(* IEC 61131-3 sources: daoli-st-library/DL_Process (part 6) *)

(* ---- FB_DL_ReactorStepCtrl.st ---- *)
(*==============================================================================
 * 组件名称 (Component)  : FB_DL_ReactorStepCtrl
 * 所属子库 (Sublibrary) : DL_Process
 * 前缀     (Prefix)     : FB_DL_
 * 当前版本 (Version)    : 1.0.1
 * 兼容性   (Platform)   : CODESYS 3.5 / TwinCAT 3 / 汇川 InoProShop / Schneider
 *                         Machine Expert；纯 IEC 61131-3（第 3 版），
 *                         仅依赖标准库 TON / R_TRIG / ABS / MAX / MIN 与库内
 *                         FB_DL_RampGenerator（IN-OUT 注入消费，斜坡不内联），
 *                         零厂商方言
 * 作者     (Author)     : 道莅代码库 · PLC编程专家（R31）
 * 开源溯源 (Origin)     : 反应釜工步顺控公开工艺语义（行业池）与 ISA-88 相
 *                         语义公开框架（暂停在步骤边界生效、恢复不重头，
 *                         主源记 T2-8），道莅 clean-room 防御性实现，
 *                         未复制任何外部源码行
 * 功能描述 (Function)   : 反应釜四工步顺控件：升温 → 保温 → 滴加 → 冷却。
 *                         温度设定经库内 FB_DL_RampGenerator 斜坡给出
 *                         （IN-OUT 注入，配方斜率单位 摄氏度每分钟 换算为
 *                         斜坡件的 摄氏度每秒 后下发）；滴加相以 bFeedAck
 *                         为终点带步超时；超温/超压独立监视层与顺控层
 *                         分离；暂停（bHold）在当前工步边界生效、恢复
 *                         不重头。不内联 PID（上层闭环外置）。
 * 复用清单 (Reuse)      : FB_DL_RampGenerator（斜坡设定，IN-OUT 注入）；
 *                         ISA-88 相语义（行为定义，零代码复制）。
 * 状态机   (States)     : eIdle/eHeat/eSoak/eFeed/eCool/eDone/ePaused/eFault，
 *                         CASE 带 ELSE 锁安全侧（fTSet 回零、停滴加）。
 * 码位     (Codes)      : 16#0005_00A8 信息级：配方域非法拒启动、配方钳位、
 *                                      暂停挂起提示（不置 bError）
 *                         16#0005_00A9 故障级：超温（独立监视层，锁存）
 *                         16#0005_00AA 故障级：超压（独立监视层，锁存）
 *                         16#0005_00AB 故障级：工步超时（滴加反馈缺失）
 *                         16#0005_00AC 故障级：状态非法（ELSE 兜底，锁存）
 * 边界防错 (Boundary)   : 1 配方域校验先于启动（斜率不大于零/温带倒置拒启动）；
 *                         2 bHold 仅在工步边界转暂停态，恢复续走原工步；
 *                         3 TON/R_TRIG 实例每拍无条件刷新；
 *                         4 CASE 带 ELSE 锁安全侧；
 *                         5 故障锁存可达解除路径：中止沿复归待机；
 *                         6 超温/超压监视独立于顺控相，任一相均生效。
 * 修订历史 (Revision)   : 2026-11-18 v1.0.0 首版入库（R31 · 阶段三 · 序 14）
 *                         2026-11-18 v1.0.1 R31 终审修复：中止/故障释放路径
 *                         补清 bError 与 uErrorId，消除释放后故障标志粘滞
 *==============================================================================*)

(*------------------------------------------------------------------------------
 * 结构体: ST_DL_ReactorRecipe（归属本功能块，同文件发布，全库唯一属主）
 *----------------------------------------------------------------------------*)
TYPE ST_DL_ReactorRecipe :
STRUCT
    fRampUp   : REAL := 2.0;    // 升温斜率 [摄氏度每分钟]，须大于 0 / Heat-up rate [degC per min], > 0
    fRampDown : REAL := 3.0;    // 降温斜率 [摄氏度每分钟]，须大于 0 / Cool-down rate [degC per min], > 0
    fSoakLo   : REAL := 80.0;   // 保温温带下限 [摄氏度] / Soak band lower [degC]
    fSoakHi   : REAL := 85.0;   // 保温温带上限 [摄氏度]，须高于下限 / Soak band upper [degC], above lower
    fFeedMl   : REAL := 50.0;   // 滴加量 [毫升] / Feed amount [mL]
    fCoolTgt  : REAL := 40.0;   // 冷却目标温度 [摄氏度] / Cool target temperature [degC]
END_STRUCT
END_TYPE

(*------------------------------------------------------------------------------
 * 枚举: E_DL_ReactorStep（归属本功能块，同文件发布，全库唯一属主）
 *----------------------------------------------------------------------------*)
TYPE E_DL_ReactorStep :
(
    eIdle   := 0,     // 待机：等待启动 / Idle, waiting for start
    eHeat   := 10,    // 升温工步：斜坡逼近温带 / Heat step, ramp to band
    eSoak   := 20,    // 保温工步：温带保持计时 / Soak step, hold band with timing
    eFeed   := 30,    // 滴加工步：等滴加反馈 / Feed step, wait feed acknowledgement
    eCool   := 40,    // 冷却工步：斜坡降到目标 / Cool step, ramp to target
    eDone   := 50,    // 完成：单拍脉冲后回待机 / Done, one-scan pulse then idle
    ePaused := 60,    // 暂停挂起：工步边界生效 / Paused, effective at step boundary
    eFault  := 99     // 故障：锁定等待中止复位 / Fault, latched until abort reset
);
END_TYPE

(*==============================================================================
 * 功能块: FB_DL_ReactorStepCtrl
 * 调用约定: 每个扫描周期无条件调用一次；ioRamp 为调用方持有的斜坡实例
 *           （IN-OUT 注入），本件驱动其引脚并读取其输出。
 *==============================================================================*)
FUNCTION_BLOCK FB_DL_ReactorStepCtrl
VAR_INPUT
    bStart   : BOOL := FALSE;         // 启动沿（待机且配方合法时受理）/ Start edge, accepted in idle with legal recipe
    bHold    : BOOL := FALSE;         // 暂停请求，工步边界生效 / Hold request, effective at step boundary
    bAbort   : BOOL := FALSE;         // 中止沿：任意态安全退出 / Abort edge, safe exit from any state
    fTNow    : REAL := 25.0;          // 釜温实测 [摄氏度] / Reactor temperature [degC]
    fPNow    : REAL := 101.0;         // 釜压实测 [千帕] / Reactor pressure [kPa]
    fPLimMax : REAL := 300.0;         // 超压监视限 [千帕]（可增引脚）/ Overpressure limit [kPa], added pin
    stRecipe : ST_DL_ReactorRecipe;   // 配方注入 / Recipe injected
    bFeedAck : BOOL := FALSE;         // 滴加完成反馈 / Feed acknowledgement feedback
    tSoak    : TIME := T#600S;        // 保温时长 [毫秒]（可增引脚）/ Soak duration [ms], added pin
    tFeedMax : TIME := T#600S;        // 滴加步超时 [毫秒]（可增引脚）/ Feed step timeout [ms], added pin
END_VAR
VAR_IN_OUT
    ioRamp   : FB_DL_RampGenerator;   // 斜坡发生器实例注入（库内复用）/ Ramp generator instance injected
END_VAR
VAR_OUTPUT
    eStep    : E_DL_ReactorStep;      // 当前工步 / Current step
    fTSet    : REAL;                  // 温度设定 [摄氏度]（斜坡输出）/ Temperature setpoint [degC]
    bFeedReq : BOOL;                  // 滴加请求 / Feed request
    bDone    : BOOL;                  // 全工步完成单拍脉冲（R27）/ All steps done one-scan pulse
    bError   : BOOL;                  // 故障标志，与故障级码配对（R45）/ Fault flag paired with fault codes
    uErrorId : UDINT;                 // 错误码，0 = 无错 / Error code, 0 = none
END_VAR
VAR
    rTrigStart: R_TRIG;               // 启动沿检测，每拍无条件刷新 / Start edge detector, refreshed every scan
    rTrigAbort: R_TRIG;               // 中止沿检测，每拍无条件刷新 / Abort edge detector, refreshed every scan
    tonSoak   : TON;                  // 保温计时，每拍无条件刷新 / Soak timer, refreshed every scan
    tonStep   : TON;                  // 步超时计时，每拍无条件刷新 / Step timeout timer, refreshed every scan
    bStepRst  : BOOL;                 // 步切换拍单拍断超时输入 / One-scan timeout break on step change
    eStatePrev: E_DL_ReactorStep;     // 上一拍步快照 / Previous step snapshot
    eResume   : E_DL_ReactorStep;     // 暂停前工步（恢复不重头）/ Step before pause, resume without restart
    bRcpOk    : BOOL;                 // 配方域合法标志 / Recipe legality flag
    bTValid   : BOOL;                 // 温度输入有效 / Temperature input validity
    bPValid   : BOOL;                 // 压力输入有效 / Pressure input validity
    bOverT    : BOOL;                 // 超温判定 / Over-temperature verdict
    bOverP    : BOOL;                 // 超压判定 / Over-pressure verdict
    uCodeLatch: UDINT;                // 故障级锁存码 / Latched fault code
    bInit     : BOOL := TRUE;         // 首扫标志 / First-scan flag
END_VAR
VAR CONSTANT
    DL_RSC_FIN   : REAL := 1.0E30;    // REAL 有限幅值判界 / REAL finiteness magnitude bound
    DL_RSC_OTMAR : REAL := 10.0;      // 超温监视裕度 [摄氏度] / Over-temp monitor margin [degC]
    DL_RSC_MIN2S : REAL := 60.0;      // 每分钟到每秒换算系数 / Per-min to per-sec factor
END_VAR

// ---- 段 1｜边沿与定时器实例无条件周期刷新（红线：禁入条件分支）----------------
rTrigStart(CLK := bStart);                            // 启动沿检测 / Start edge detection
rTrigAbort(CLK := bAbort);                            // 中止沿检测 / Abort edge detection
tonSoak(IN := (eStep = eSoak) AND (NOT bHold), PT := tSoak); // 保温计时，暂停断输入 / Soak timing, broken on hold
tonStep(IN := (eStep = eFeed) AND (NOT bStepRst), PT := tFeedMax); // 滴加超时按步断输入 / Feed timeout per step

// ---- 段 2｜步切换检测 ------------------------------------------------------------
bStepRst := (eStep <> eStatePrev) OR bInit;           // 步变化即断输入 / Step change breaks timing
eStatePrev := eStep;                                  // 快照留痕 / Snapshot previous step
bInit := FALSE;                                       // 清首扫标志 / Clear first-scan flag

// ---- 段 3｜输入有效性与独立监视层判定（与顺控相分离）------------------------------
bTValid := (fTNow = fTNow) AND (ABS(fTNow) < DL_RSC_FIN);   // 温度有限 / Temperature finite
bPValid := (fPNow = fPNow) AND (ABS(fPNow) < DL_RSC_FIN);   // 压力有限 / Pressure finite
bOverT  := bTValid AND (eStep <> eIdle) AND (fTNow > stRecipe.fSoakHi + DL_RSC_OTMAR); // 超温：带外裕度判 / Over-temp beyond margin
bOverP  := bPValid AND (eStep <> eIdle) AND (fPNow > fPLimMax); // 超压独立判 / Over-pressure independent
IF bOverT THEN
    uCodeLatch := 16#0005_00A9;                       // 码位：超温 / Code: over temperature
END_IF
IF bOverP THEN
    uCodeLatch := 16#0005_00AA;                       // 码位：超压 / Code: over pressure
END_IF
IF bOverT OR bOverP THEN
    eStep := eFault;                                  // 监视层直接锁故障 / Monitor layer latches fault directly
END_IF

// ---- 段 4｜中止沿统一入口：停滴加、温度设定回零、复归待机 ------------------------
IF rTrigAbort.Q THEN
    eStep := eIdle;                                   // 中止复归待机 / Abort returns to idle
    bFeedReq := FALSE;                                // 停滴加请求 / Stop feed request
    bError := FALSE;                                  // 中止含故障态释放路径，清故障标志（R28 终审）/ Abort is fault release path, clears flag
    uErrorId := 16#0000_0000;                         // 中止清错误码防粘滞（R28 终审）/ Abort clears error code against stickiness
END_IF

// ---- 段 5｜状态机（CASE 带 ELSE 锁安全侧：fTSet 回零、停滴加）---------------------
CASE eStep OF
    eIdle:
        fTSet := 0.0;                                 // 待机设定回零（安全侧）/ Idle setpoint zero, safe side
        bFeedReq := FALSE;                            // 待机停滴加 / Idle stops feed
        bDone := FALSE;                               // 清完成脉冲 / Clear done pulse
        ioRamp(bEnable := FALSE, bTrack := TRUE, fTrackValue := fTNow); // 斜坡跟踪实测免扰动 / Ramp tracks actual
        IF rTrigStart.Q THEN
            bRcpOk := (stRecipe.fRampUp > 0.0) AND (stRecipe.fRampDown > 0.0)
                  AND (stRecipe.fSoakLo < stRecipe.fSoakHi)
                  AND (stRecipe.fFeedMl >= 0.0) AND (stRecipe.fCoolTgt < stRecipe.fSoakLo)
                  AND (stRecipe.fRampUp < DL_RSC_FIN) AND (stRecipe.fRampDown < DL_RSC_FIN); // 配方域校验先于启动 / Recipe check before start
            IF bRcpOk THEN
                eStep := eHeat;                       // 配方合法进升温 / Legal recipe, to heat
            ELSE
                uErrorId := 16#0005_00A8;             // 信息级：配方非法拒启动 / Info: illegal recipe, start rejected
            END_IF
        END_IF
    eHeat:
        bFeedReq := FALSE;                            // 升温停滴加 / Heat stops feed
        ioRamp(bEnable := TRUE, fTarget := stRecipe.fSoakHi,
               fRateUp := stRecipe.fRampUp / DL_RSC_MIN2S,
               fRateDown := stRecipe.fRampDown / DL_RSC_MIN2S,
               bHold := FALSE);                       // 斜坡下发，配方斜率换算每秒 / Ramp driven, rate per second
        fTSet := ioRamp.fOut;                         // 温度设定取斜坡输出 / Setpoint from ramp output
        IF ioRamp.bDone AND bTValid AND (fTNow >= stRecipe.fSoakLo) THEN
            eStep := eSoak;                           // 到带复验后转保温（R42）/ Recheck then to soak
        END_IF
        IF bHold AND ioRamp.bDone THEN
            eResume := eSoak;                         // 边界暂停登记续点（ISA-88）/ Boundary pause books resume step
            eStep := ePaused;                         // 转暂停挂起 / To paused
        END_IF
    eSoak:
        bFeedReq := FALSE;                            // 保温停滴加 / Soak stops feed
        ioRamp(bEnable := TRUE, fTarget := stRecipe.fSoakHi,
               fRateUp := stRecipe.fRampUp / DL_RSC_MIN2S,
               fRateDown := stRecipe.fRampDown / DL_RSC_MIN2S,
               bHold := FALSE);                       // 保温维持带顶设定 / Soak holds band top
        fTSet := ioRamp.fOut;                         // 温度设定取斜坡输出 / Setpoint from ramp output
        IF tonSoak.Q THEN
            eStep := eFeed;                           // 保温满转滴加 / Soak elapsed, to feed
        END_IF
        IF bHold THEN
            eResume := eSoak;                         // 边界暂停登记续点 / Boundary pause books resume step
            eStep := ePaused;                         // 转暂停挂起 / To paused
        END_IF
    eFeed:
        bFeedReq := TRUE;                             // 滴加请求置位 / Feed request set
        fTSet := ioRamp.fOut;                         // 温度设定维持 / Setpoint maintained
        IF tonStep.Q THEN
            eStep := eFault;                          // 滴加反馈缺失锁故障（步超时）/ Feed ack missing, fault
            uCodeLatch := 16#0005_00AB;               // 码位：步超时/反馈缺失 / Code: step timeout
        ELSIF bFeedAck THEN
            eStep := eCool;                           // 滴加完成转冷却 / Feed done, to cool
        END_IF
    eCool:
        bFeedReq := FALSE;                            // 冷却停滴加 / Cool stops feed
        ioRamp(bEnable := TRUE, fTarget := stRecipe.fCoolTgt,
               fRateUp := stRecipe.fRampUp / DL_RSC_MIN2S,
               fRateDown := stRecipe.fRampDown / DL_RSC_MIN2S,
               bHold := FALSE);                       // 斜坡降到冷却目标 / Ramp down to cool target
        fTSet := ioRamp.fOut;                         // 温度设定取斜坡输出 / Setpoint from ramp output
        IF ioRamp.bDone AND bTValid AND (fTNow <= stRecipe.fCoolTgt + 1.0) THEN
            eStep := eDone;                           // 到目标复验后转完成（R42）/ Recheck then to done
        END_IF
        IF bHold AND ioRamp.bDone THEN
            eResume := eDone;                         // 边界暂停登记续点 / Boundary pause books resume step
            eStep := ePaused;                         // 转暂停挂起 / To paused
        END_IF
    eDone:
        fTSet := ioRamp.fOut;                         // 完成态维持设定 / Done maintains setpoint
        bFeedReq := FALSE;                            // 完成停滴加 / Done stops feed
        bDone := TRUE;                                // 完成单拍脉冲 / One-scan done pulse
        eStep := eIdle;                               // 下拍回待机 / Back to idle next scan
    ePaused:
        fTSet := ioRamp.fOut;                         // 暂停冻结设定（斜坡 bHold 语义由态承载）/ Pause freezes setpoint
        bFeedReq := FALSE;                            // 暂停停滴加 / Pause stops feed
        uErrorId := 16#0005_00A8;                     // 信息级：暂停挂起提示 / Info: paused notice
        IF (NOT bHold) AND (eResume <> ePaused) THEN
            eStep := eResume;                         // 恢复不重头续走原工步 / Resume without restart
        END_IF
    eFault:
        fTSet := 0.0;                                 // 故障安全侧设定回零 / Fault safe side setpoint zero
        bFeedReq := FALSE;                            // 故障停滴加 / Fault stops feed
        bDone := FALSE;                               // 故障清完成 / Fault clears done
        IF rTrigAbort.Q THEN
            eStep := eIdle;                           // 可达解除路径：中止沿复归 / Reachable release: abort edge
            uCodeLatch := 16#0000_0000;               // 清锁存码 / Clear latched code
            bError := FALSE;                          // 释放同步清故障标志（R28 终审）/ Release clears fault flag
            uErrorId := 16#0000_0000;                 // 释放同步清错误码 / Release clears error code
        END_IF
    ELSE
        eStep := eFault;                              // 非法状态兜底 / Illegal state fallback
        uCodeLatch := 16#0005_00AC;                   // 码位：状态非法 / Code: illegal state
        fTSet := 0.0;                                 // 兜底设定回零（安全侧）/ Fallback setpoint zero
        bFeedReq := FALSE;                            // 兜底停滴加 / Fallback stops feed
END_CASE

// ---- 段 6｜错误码装配：故障锁存回放优先，信息级居次 ------------------------------
IF eStep = eFault THEN
    bError   := TRUE;                                 // 故障标志配对（R45）/ Fault flag paired
    uErrorId := uCodeLatch;                           // 故障码锁存回放 / Latched fault code replayed
END_IF
END_FUNCTION_BLOCK

(* ---- FB_DL_ReworkLotGate.st ---- *)
(*
  ==================================================================
  组件名 Component  : FB_DL_ReworkLotGate
  分类   Category   : DL_Process
  前缀   Naming     : FB_DL_ ｜ b/n/u/f/t/e/st 类型前缀制（R265）
  码位   Code ID    : 16#0006_3036（故障级：越权放行锁存）｜ 16#0006_3037
                      （信息级：放行计数饱和钳位）
  版本   Version    : 1.0.1
  变更   CHANGELOG  : v1.0.1 eReleased 放行相单拍回迁
  复杂度 Complexity  : 中
  功能   Purpose    : 返工批拦截闸：返工标记登记期拦截放行指令，复检合格才
                      放行并计数；返工登记期未复检合格的放行指令判「越权
                      放行」并锁存故障；供批次放行合规审计与质量门禁使用。
  开源溯源 Origin    : ISA-88 批次相状态模型（公开条款，R12 沿用）+ PackML
                      纪律次源（T2-7 / T2-8）：仅借「批次相语义」状态命名
                      组织方式；返工闸逻辑完全自研，零代码复制。
  许可证 License    : MIT
  参考   Reference  : IEC 61131-3:2013 §6.6 状态机 / R_TRIG 语义；ISA-88
                      批次相状态公开条款（借语义，不抄文）
  平台   Platform   : 纯 IEC 61131-3（R_TRIG / ENUM+CASE / 四则），三平台通用
  依赖   Depends    : 仅 Standard.library（R_TRIG 属标准件）
  分工声明 Split     : FB_DL_BatchPhaseTrack（批次相跟踪）/ FB_DL_HoldResumeSeq
                      （保持恢复顺控）与本件互引；本件只管「返工标记 → 放行
                      合规」单门禁，不做批次全程跟踪（R216）。
  归属 Ownership     : E_DL_ReworkGatePhase 属主为本文件（全库唯一定义，R264）；
                      引用件只引用不重声明。
  ------------------------------------------------------------------
  边界 Boundary     :
                      一 组态口径（定稿，R90 反证句见码表）：nQuotaMax < 1
                         按「钳位接管为 1」静默接管——上限为 1 的闸仍有
                         完整拦截语义（登记 + 复检合格才放行 + 计数），
                         功能不静默丢失，非永假防御；不为此另立故障码
                         （组态缺省出口与正常运行出口完全同形：闸照常
                         工作、计数照常推进，无任何输出可区分该场景）；
                         3036 专用于越权放行锁存；
                      二 状态机 ENUM + CASE 必带 ELSE（非法态兜底落 eFault +
                         锁存 3036，禁静默）；本拍合法事件（复检合格沿 /
                         登记撤除）优先于越权判据（R275 同拍竞态）；
                      三 越权放行判据（锁存回放，R152）：返工登记电平 +
                         放行指令 + 复检未合格 → 锁存 3036 + bError；
                         锁存解除式（可达自证）：bResetCmd 上升沿清锁存
                         回 eIdle（输入引脚恒可达，无「置位即永久」路径）；
                      四 合规放行计数：放行沿（rtRelease R_TRIG，段 0 无条件
                         刷新）+ 复检合格 + 未锁存才计数；计数达 nQuotaMax
                         饱和钳位 + 信息级 3037（不置 bError，闸功能不受
                         影响，钳位为审计口径不是功能门槛）；
                      五 bEnable = FALSE 的语义写死（FB33-4 声明行）：强制
                         eIdle + 双出口复位（不 faults，使能断开 ≠ 合规故障）；
                      六 首拍 _bInit 全量初始化；无浮点量、无除法、无定时器
                         （纯电平 / 沿 / 计数语义）；无全局、无外部变量、
                         无物理地址。
  错误码 Codes      :
    16#0006_3036【故障级】越权放行（返工登记期放行指令且复检未合格）或非法
                         状态拦截（ELSE 兜底），锁存回放至复位沿
    16#0006_3037【信息级】放行计数已达 nQuotaMax 饱和钳位（不置 bError）
  码位反证 Note     :
    3036 与 3037 不可合并：3036 锁存 + bValid = FALSE + bError = TRUE，
    3037 不锁存 + bValid = TRUE + bError = FALSE，bValid / bError 双通道
    可唯一区分，按 R90 分立；「登记撤除瞬间的放行沿」与「越权」由同拍
    事件优先序区分（边界二），不需第三码。
  验收 Acceptance   :
    算法已证（脚本）：未跑 ｜ 编译器已证（三平台）：未跑
    V1 无登记 + 放行沿 → nReleased + 1、bReleaseAllow（正常批口径）
    V2 登记 + 复检合格 + 放行沿 → 计数 + 1（返工批合规放行）
    V3 登记 + 复检未合格 + 放行指令 → 锁存 3036 + bError
    V4 锁存态 bResetCmd 上升沿 → 解锁回 eIdle（锁存解除可达向量）
    V5 nQuotaMax = 3、放行 4 次 → nReleased 钳 3 + 码 3037
       （bError = FALSE，闸功能照常）
    V6 nQuotaMax = 0 → 钳位接管为 1（边界一定稿口径，功能不静默丢失）
    V7 失能 → eIdle + 双出口复位（不 faults）
    V8 非法枚举态（强改 eState）→ ELSE 兜底落 eFault + 3036
  修订记录 Revision  :
    2026-11-21  v1.0.0  R64 首版（批 3 · 序号 9，ISA-88 / PackML 纪律次源 + 自研）
    2026-11-22  v1.0.1  R65 点修（eReleased 回迁，R64 终审项）：v1.0.0 放行相
                        在 bReleaseCmd 持续保持且无再登记时停留该相不回迁，
                        下批次无法进入；v1.0.1 改放行相为单拍驻留相——完成后
                        无条件回迁待判 / 空闲相 eIdle；回迁清理声明：本件无
                        放行锁存与批次暂存变量（rtRelease 为自清沿实例，
                        Q 单拍自灭；nReleased 为审计台账不属暂存，复位沿亦
                        不清，边界四口径），回迁即天然清零，无需额外清零动作；
                        登记电平若仍生效，由 eIdle 相在下一拍重新迁入拦截相
                        （合法重入，rtRelease 沿不自触发，计数不受影响）
  ==================================================================
*)
TYPE E_DL_ReworkGatePhase :
(
    eIdle       := 0,  // 待机：无返工登记 / idle, no rework registered
    eReworkHold := 10, // 返工拦截：登记生效，等复检合格 / the rework hold, waiting for the recheck pass
    eReleased   := 20, // 放行：合规放行相（登记撤除或复检合格放行后驻留一拍语义由调用方承接）/ the released phase
    eFault      := 30  // 锁存故障：越权放行或非法态，复位沿解除 / a latched fault released by the reset edge
);
END_TYPE

FUNCTION_BLOCK FB_DL_ReworkLotGate
VAR_INPUT
    bEnable      : BOOL := TRUE;  // 使能，FALSE 时强制 eIdle + 双出口复位（边界五）/ the enable, false forces the idle and resets both outlets
    bLotRework   : BOOL := FALSE; // 返工标记登记电平 [-]（来自批次履历）/ the rework registration level from the lot history
    bRecheckPass : BOOL := FALSE; // 复检合格电平 [-] / the recheck pass level
    bReleaseCmd  : BOOL := FALSE; // 放行指令电平 [-] / the release command level
    bResetCmd    : BOOL := FALSE; // 故障复位电平，上升沿清锁存回 eIdle（边界三解除式）/ the fault reset level, its rising edge releases the latch
    nQuotaMax    : DINT  := 16;   // 放行计数饱和上限 [个]，须 ≥ 1，< 1 钳位接管为 1（边界一定稿）/ the release count ceiling, at least one, clamped when below
END_VAR
VAR_OUTPUT
    bReleaseAllow : BOOL := FALSE;           // 放行许可电平 [-]（锁存 / 失能强制 FALSE）/ the release permission forced false on a latch or disable
    bReworkHold   : BOOL := FALSE;           // 返工拦截中指示 [-] / the rework hold indicator
    nReleased     : DINT  := 0;              // 合规放行计数 [个]（饱和口径）/ the compliant release count saturated
    eState        : E_DL_ReworkGatePhase;    // 状态机出口 [状态] / the state machine outlet
    bValid        : BOOL := FALSE;           // 判据可用 [-] / the criteria are usable
    eErr          : UDINT := 16#0000_0000;   // 错误码，0 = 正常 / the error code, zero is ok
    bError        : BOOL := FALSE;           // 故障标志（故障级码同拍置位，R45 配对）/ the fault flag raised with a fault level code
END_VAR
VAR
    _bInit      : BOOL := FALSE;  // 首拍初始化标志（R310 / FB50-2）/ the first scan flag
    _eState     : E_DL_ReworkGatePhase := E_DL_ReworkGatePhase.eIdle; // 内部状态寄存器 / the internal state register
    _bFaultLatch: BOOL := FALSE;  // 故障锁存副本（仅复位沿清除）/ the fault latch copy
    _uLatch     : UDINT := 16#0000_0000; // 故障码锁存 [码]（复位沿清除，FB33-1）/ the latched fault code cleared by the reset edge
    _nReleased  : DINT  := 0;     // 计数内部副本 [个]（饱和钳位口径）/ the internal count copy saturated
    _nQuotaUse  : DINT  := 1;     // 上限接管量 [个]（< 1 钳位为 1，边界一）/ the ceiling taken over clamped to one
    _bCountSat  : BOOL := FALSE;  // 计数饱和标记（单拍信息位，段 6 映射）/ the count saturation flag of this scan
    rtReset     : R_TRIG;         // 复位沿实例，段 0 无条件刷新（R7）/ the reset edge instance refreshed unconditionally
    rtRelease   : R_TRIG;         // 合规放行沿实例，段 0 无条件刷新 / the compliant release edge instance refreshed unconditionally
END_VAR  // R64 结构补齐：VAR 段缺失的 END_VAR（门禁机械修复）
VAR CONSTANT
    DL_RLG_ZEROI: DINT  := 0;  // 整型零常量 [个] / the integer zero constant
    DL_RLG_ONEI : DINT  := 1;  // 整型一常量 [个] / the integer one constant
    DL_RLG_ZEROU: UDINT := 16#0000_0000; // 码零常量 / the code zero constant
END_VAR

// 段 0｜沿检测无条件周期刷新（禁入分支，R7）/ segment 0, the unconditional edge refresh
rtReset(CLK := bResetCmd); // 复位沿 / the reset edge
rtRelease(CLK := bReleaseCmd AND NOT _bFaultLatch AND bEnable
                 AND (NOT bLotRework OR bRecheckPass)); // 合规放行沿（登记撤除或复检合格的放行指令上升沿，R275 事件优先口径）/ the compliant release edge of the legal command

// 段 1｜首拍初始化与复位沿作用域（R310 / R311）/ segment 1, the first scan init and the reset edge scope
IF NOT _bInit THEN // 首拍一拍 / the first scan
    _bInit := TRUE; // 置首拍标志 / raise the first scan flag
    _eState := E_DL_ReworkGatePhase.eIdle; // 状态显式落空闲 / place the state to idle
    _bFaultLatch := FALSE; // 故障锁存显式清零 / clear the fault latch explicitly
    _uLatch := DL_RLG_ZEROU; // 码锁存显式清零 / clear the latched code explicitly
    _nReleased := DL_RLG_ZEROI; // 计数显式清零 [个] / clear the count explicitly
    _nQuotaUse := DL_RLG_ONEI; // 上限接管显式置一 [个] / preset the ceiling one explicitly
END_IF
IF rtReset.Q THEN // 复位沿（作用域声明：清锁存 + 迁相位，不清计数——计数是审计台账，R311）/ the reset edge with the declared scope, the audit count survives
    _bFaultLatch := FALSE; // 清故障锁存（唯一解除路径，边界三自证可达）/ clear the fault latch, the only release path
    _uLatch := DL_RLG_ZEROU; // 清码锁存 / clear the latched code
    _eState := E_DL_ReworkGatePhase.eIdle; // 迁回空闲 / back to idle
END_IF

// 段 2｜上限接管与计数饱和预置（边界一：nQuotaMax < 1 钳位接管为 1，功能不静默丢失）/ segment 2, the ceiling take over and the saturation preset
_nQuotaUse := nQuotaMax; // 上限接管 [个] / take the ceiling
IF _nQuotaUse < DL_RLG_ONEI THEN // 上限 < 1（组态缺省）/ the ceiling below one
    _nQuotaUse := DL_RLG_ONEI; // 钳位接管为 1（拦截闸仍有完整语义）/ clamp to one, the gate keeps its full semantics
END_IF
_bCountSat := FALSE; // 计数饱和标记预清零（单拍信息位，R256 统一出口预置）/ preset the saturation flag false

// 段 3｜失能分支：强制 eIdle + 双出口复位，不 faults（边界五声明行）/ segment 3, the disabled branch
IF NOT bEnable THEN // 失能 / disabled
    _eState := E_DL_ReworkGatePhase.eIdle; // 强制空闲 / force the idle
    _bFaultLatch := FALSE; // 锁存复位（使能断开 ≠ 合规故障）/ clear the latch
    _uLatch := DL_RLG_ZEROU; // 码锁存复位 / clear the code
    eState := _eState; // 状态出口 / the state outlet
    bReleaseAllow := FALSE; // 许可电平复位 / the permission resets
    bReworkHold := FALSE; // 拦截指示复位 / the hold indicator resets
    bValid := FALSE; // 失能即不可用 / the criteria are not usable while disabled
    bError := FALSE; // 失能不是故障 / a disabled device is not a fault
    eErr := DL_RLG_ZEROU; // 失能不发码 / no code is emitted while disabled
    RETURN; // 早退（计数不动，失能不清审计台账）/ early return, the audit count survives
END_IF

// 段 4｜主状态机（ENUM + CASE，ELSE 兜底；本拍事件优先于越权判据，R275）/ segment 4, the main machine, the event before the misuse verdict
CASE _eState OF
    E_DL_ReworkGatePhase.eIdle: // 空闲相 / the idle phase
        IF bLotRework THEN // 返工登记生效 / the rework registration is active
            _eState := E_DL_ReworkGatePhase.eReworkHold; // 迁入拦截相 / enter the hold phase
        END_IF
    E_DL_ReworkGatePhase.eReworkHold: // 返工拦截相（本拍合法事件优先：登记撤除或复检合格放行先消化，再消化越权判据，R275）/ the hold phase, the legal event before the misuse
        IF NOT bLotRework THEN // 事件优先：登记撤除 / the registration withdrawn, the event goes first
            _eState := E_DL_ReworkGatePhase.eIdle; // 回空闲 / back to idle
        ELSIF bRecheckPass AND bReleaseCmd THEN // 复检合格 + 放行指令（合规放行，边界四口径）/ the recheck passed with the release command
            _eState := E_DL_ReworkGatePhase.eReleased; // 迁入放行相 / enter the released phase
        ELSIF bReleaseCmd THEN // 越权判据：登记中放行且复检未合格（真实可达：操作员越过复检直接放令）/ the misuse path, reachable by the operator bypassing the recheck
            _bFaultLatch := TRUE; // 锁存故障 / latch the fault
            _uLatch := 16#0006_3036; // 故障级：越权放行 / fault grade, the unauthorized release
            bError := TRUE; // 同拍置故障标志（R45 配对，段 6 故障分支沿用）/ raise the fault flag on the same scan
        END_IF
    E_DL_ReworkGatePhase.eReleased: // 放行相（v1.0.1 改单拍驻留：完成后强制回迁空闲，R64 终审修复「eReleased 不回迁」）/ the released phase, single scan dwell with the forced return since v1.0.1
        _eState := E_DL_ReworkGatePhase.eIdle; // 放行相完成后无条件回迁待判 / 空闲相（下批次可正常进入；v1.0.0 在 bReleaseCmd 持续保持且无再登记时停留该相不回迁，为本次修复点）/ unconditional return to idle after the release completes
        // 回迁清理声明（v1.0.1）：本件无放行锁存与批次暂存变量——rtRelease 为自清沿实例（Q 单拍自灭），nReleased 为审计台账不属暂存（复位沿亦不清，边界四），回迁即天然清零，无额外清零动作 / no release latch or batch staging exists, the return clears naturally
    E_DL_ReworkGatePhase.eFault: // 锁存故障相（驻留，解除由段 1 复位沿承担）/ the fault phase dwelling, the release belongs to the reset edge
        ; // 驻留语义由注释表达（禁自赋值死语句，R261）/ the dwell is expressed by this comment without a dead statement
    ELSE // 非法枚举值拦截（边界二：落故障相并锁存，禁静默）/ the illegal enumeration guard
        _bFaultLatch := TRUE; // 锁存故障 / latch the fault
        _uLatch := 16#0006_3036; // 故障级：非法状态拦截（归入越权族一码，出口同形锁存回放，R90）/ fault grade, the illegal state under the latch family
        bError := TRUE; // 同拍置故障标志（R45 配对）/ raise the fault flag on the same scan
        _eState := E_DL_ReworkGatePhase.eFault; // 落故障相 / force the fault phase
END_CASE

// 段 5｜合规放行计数（边界四：沿 + 未锁存才计数；饱和钳位 + 信息级）/ segment 5, the compliant release counting with the saturation
IF rtRelease.Q AND (NOT _bFaultLatch) THEN // 合规放行沿且未锁存 / a compliant release edge without a latch
    IF _nReleased < _nQuotaUse THEN // 计数未达上限 / the count below the ceiling
        _nReleased := _nReleased + DL_RLG_ONEI; // 计数推进 [个] / advance the count
    ELSE // 计数已达上限：饱和钳位 + 信息级（闸功能不受影响，边界四）/ the count saturated with the info code, the gate unaffected
        _bCountSat := TRUE; // 置饱和标记（单拍信息位）/ raise the saturation flag
    END_IF
END_IF

// 段 6｜故障锁存迁移闸 + 统一出口（名实双出口同源，R191）/ segment 6, the latch gate and the unified outlet
IF _bFaultLatch AND (_eState <> E_DL_ReworkGatePhase.eFault) THEN // 已锁存但不在故障相 / latched outside the fault phase
    _eState := E_DL_ReworkGatePhase.eFault; // 迁入故障相 / enter the fault phase
END_IF
eState := _eState; // 状态出口 / the state outlet
bReleaseAllow := (NOT _bFaultLatch) AND bEnable
              AND ((NOT bLotRework) OR bRecheckPass); // 许可电平与判据同源派生（登记中须复检合格）/ the permission derived from the criteria
bReworkHold := (_eState = E_DL_ReworkGatePhase.eReworkHold); // 拦截指示与状态同源 / the hold indicator from the state
nReleased := _nReleased; // 计数出口 [个] / the count outlet
IF _bFaultLatch THEN // 故障锁存回放优先（不在故障相按当下输入重新推断，R152）/ the latched fault replays first
    bValid := FALSE; // 故障相不可用 / not usable in the fault phase
    bError := TRUE; // 故障位置位（R45 配对）/ raise the fault bit
    eErr := _uLatch; // 锁存码回放 / replay the latched code
ELSIF _bCountSat THEN // 计数饱和（信息级，单拍重算）/ the saturation, informational
    bValid := TRUE; // 闸功能照常可用 / the gate stays usable
    bError := FALSE; // 信息级不置故障标志（R285）/ keep the fault flag false
    eErr := 16#0006_3037; // 信息级：放行计数饱和钳位 / informational, the count saturated
ELSE // 无事件 / no event
    bValid := TRUE; // 判据可用 / the criteria are usable
    bError := FALSE; // 无故障 / no fault
    eErr := DL_RLG_ZEROU; // 正常 / ok
END_IF
END_FUNCTION_BLOCK

(* ---- FB_DL_RotaryIndexTable.st ---- *)
(*==============================================================================
 * 组件名称 (Component)  : FB_DL_RotaryIndexTable
 * 所属子库 (Sublibrary) : DL_Process
 * 当前版本 (Version)    : 1.0.0
 * 组件分类 (Category)   : 功能块（FUNCTION_BLOCK）· 工站模板 · 多工位分度盘调度
 * 兼容性 (Platform)     : CODESYS 3.5 / TwinCAT 3 / 汇川 InoProShop / Machine Expert；
 *                         仅依赖标准库（TON / R_TRIG / F_TRIG / LIMIT），分度请求
 *                         以布尔脉冲出口下发，块内不绑定任何电机或驱动库
 * 功能描述 (Function)   : 管理「分度请求 → 到位确认 → 稳定等待 → 工位工艺放行」的
 *                         节拍链；维护工位启用表与工艺号映射，支持空跑（清洗）模式
 *                         逐位走完，并对分度超时与到位信号抖动给出可诊断的故障码
 * 与既有件边界 (Scope)  : 料仓槽位台账（空 / 满 / 不合格）由料仓件承担，本块不管槽
 *                         位内容；连续输送积放由输送段件承担，本块管离散分度盘的节
 *                         拍与工位放行。三者拓扑互斥，语义不重叠
 * 状态机规模 (States)   : 五态最小子集（eIdle 0 / eDwell 10 / eIndexing 20 /
 *                         eSettling 30 / eFault 99）。eSettling 单独成态，用于隔离
 *                         「到位后抖动」的诊断窗口，避免把机械抖动混入分度超时计数
 * 关键算法 (Algorithm)  :
 *   ① 工位号合法性：nAtStation 须落在 1~生效工位数，越界即 02D2，不做猜测性修正
 *   ② 掩码构造：每拍由启用表重建，逐位置位（位累加器左移一位再或），不拼累计量，
 *      规避位宽边界；工位数上限 24，恒在安全域内
 *   ③ 停留计时：剩余停留时间由定时器已历时反算，空跑模式直接旁路计时
 *   ④ 空跑模式：工艺放行恒假，分度链照走，用于清洗与调试；不计循环数
 *   ⑤ 循环计数：分度回到 1 号位那一拍出单拍脉冲并累加，饱和防溢出
 *   ⑥ 抖动诊断：稳定窗内到位信号掉沿即判硬件问题，直接锁故障且不自动重试——自动
 *      重试会把机械松动掩盖成偶发超时，现场极难定位
 * 码位表 (Error codes)  :
 *   16#0005_01C2【信息级】工位数量越界已钳位至 2~24，不置故障位
 *   16#0005_02D0【故障级】分度超时（到位信号未在监控窗内建立）
 *   16#0005_02D1【故障级】到位信号抖动或丢失（稳定窗内掉沿）
 *   16#0005_02D2【故障级】工位号越界（机械到位反馈不可信）
 *   16#0005_02D3【故障级】非法状态兜底
 * R32 写入点次序审计 :
 *   nActiveStation  : ① 空跑 / 停机撤销时清 0（段 6、段 7）→ ② 停留与稳定段按到位
 *                     反馈刷新（eDwell / eSettling 各一处，同拍只可能命中一处）
 *   bStationReady   : 仅段 10 单点派生（由生效工位数、启用表、空跑模式三者与门），
 *                     状态机内不写，杜绝分支双写
 *   nRecipeAtStation: 仅段 10 单点派生（工艺号透传，越界给 0，不做校验）
 *   tDwellRemain    : 仅段 10 单点派生（由停留定时器已历时反算，钳位非负）
 *   _uErrorIdInt    : ① 首扫清（段 4）→ ② 分度超时（eIndexing）→ ③ 抖动（eSettling）
 *                     → ④ 工位号越界（eSettling）→ ⑤ 非法状态（ELSE）→ ⑥ 复位清
 *   _eState         : 每拍只在 CASE 分支出口单点写入；CASE 之外仅段 6 使能撤销一处
 * 设计偏离登记 (Deviations) :
 *   D1 增补 tCycle 引脚（默认 10 毫秒）：统计结构体内含累计运行时长，而块内无时间
 *      基准引脚则无法累加；按库内既有公约以任务扫描周期作基准，向后兼容（有默认
 *      值），不改变任何既有引脚语义
 *   D2 分度计数在「到位确认通过」拍累加，而非请求拍：超时未到位属失败分度，不应
 *      计入成功次数；与规格文字「分度次数」取成功口径一致
 * 验收向量 (Acceptance) :
 *   V1 掩码：工位数 8、前 5 个启用 → 掩码 16#0000_001F
 *   V2 工艺号透传：到位 3 号工位、3 号工艺号 27 → 作业工位 3、工艺号 27、放行为真
 *   V3 分度超时：监控窗 2 秒内到位信号未建立 → 码 02D0、故障态、故障位为真
 *   V4 空跑：工位数 4、空跑为真 → 逐位推进，4 拍后出循环脉冲，循环计数不增
 *   V5 抖动：到位后 50 毫秒内信号由真转假 → 码 02D1，无自动重试
 * 开源溯源 (Origin)     : 参考包装机械公开手册的工位 / 节拍语义组织与位掩码工位表
 *                         写法，只借分类与参数域；状态机、掩码重建、抖动诊断、码位
 *                         与引脚契约为本库独立设计，clean-room 不构成衍生作品
 * 红线自检 (Redline)    : R1 零全局表与外部变量引用、零物理地址记号 ✓｜R2 零占位符 ✓
 *                         R3 纯 IEC 61131-3 加标准库 ✓｜R4 数组先判界、除法防零、
 *                         时长反算钳非负 ✓｜R5 声明行中英双语同行注释 ✓｜R6 五成员逐
 *                         一有 CASE 标签且含 ELSE 兜底 ✓｜R7 三沿检测（启动 / 停止 /
 *                         复位）与到位双沿、三定时器全部在 CASE 之外无条件刷新 ✓
 * 修订历史 (Revision)   :
 *   2026-11-15  v1.0.0  首版入库（Round 11 · C 泳道 · 工站四件套之二）
 *============================================================================*)

(*------------------------------------------------------------------------------
 * 枚举: E_DL_IndexTableState（归属 FB_DL_RotaryIndexTable，同文件发布）
 *   五态，每个成员在主状态机中均有同名 CASE 标签（R31 完备性）
 *-----------------------------------------------------------------------------*)
TYPE E_DL_IndexTableState :
(
    eIdle     := 0,     // 待机：等启动沿，不发放行 / Idle, awaiting start, no permit
    eDwell    := 10,    // 停留：当前工位工艺放行窗 / Dwell, process permit window
    eIndexing := 20,    // 分度中：已出请求脉冲，等到位 / Indexing, waiting for in-position
    eSettling := 30,    // 稳定中：到位后去抖确认 / Settling, debounce after in-position
    eFault    := 99     // 故障锁存：仅复位沿可退 / Fault latched, only a reset edge leaves
);
END_TYPE

(*------------------------------------------------------------------------------
 * 结构体: ST_DL_IndexTableStat（归属 FB_DL_RotaryIndexTable）
 *   跨周期统计，由调用方持有，本块只累加，掉电保持由上层负责
 *-----------------------------------------------------------------------------*)
TYPE ST_DL_IndexTableStat :
STRUCT
    nIndexCount : UDINT;                    // 累计成功分度次数 [次] [Successful index counter]
    nCycleCount : UDINT;                    // 累计整圈循环数 [圈] [Full revolution counter]
    tRunTime    : TIME;                     // 累计运行时长 [毫秒] [Accumulated run time]
END_STRUCT
END_TYPE

FUNCTION_BLOCK FB_DL_RotaryIndexTable
VAR_INPUT
    bEnable          : BOOL;                            // 使能，FALSE 撤销分度请求并回待机 [Enable, withdraws request on FALSE]
    bStart           : BOOL;                            // 启动节拍循环，上升沿受理 [Start the cycle on a rising edge]
    bStop            : BOOL;                            // 完成当前工位后停止，上升沿受理 [Stop after current station, rising edge]
    bReset           : BOOL;                            // 复位故障，上升沿受理 [Reset fault on rising edge]
    nStationCount    : INT;                             // 工位总数 [个]，有效域 2~24 [Station count, 2..24]
    nAtStation       : INT;                             // 机械到位工位号 [1~工位数]，0 表示未定位 [Mechanical station number, 0 = not seated]
    bIndexInPos      : BOOL;                            // 分度到位开关信号 [-] [Indexer in-position switch]
    abStationEnable  : ARRAY[1..24] OF BOOL;            // 工位启用表，FALSE 视为空位 [Station enable table, FALSE = empty]
    anStationRecipe  : ARRAY[1..24] OF INT;             // 工位工艺号表，仅透传不校验 [-] [Per-station recipe number, pass-through]
    tDwellTime       : TIME := T#1S;                    // 每工位停留时间 [毫秒]，0 表示不停留 [Dwell per station]
    tSettleTime      : TIME := T#100MS;                 // 到位后稳定确认时间 [毫秒]，滤机械抖动 [Settling time after in-position]
    tIndexTimeout    : TIME := T#3S;                    // 分度超时 [毫秒]，0 表示不监控 [Indexing timeout]
    bDryRun          : BOOL;                            // 空跑（清洗）模式：忽略启用表逐位走完 [Dry-run mode, ignores enable table]
    tCycle           : TIME := T#10MS;                  // 任务扫描周期 [毫秒]，累计运行时长基准（偏离 D1）[Task cycle time, run-time base]
END_VAR
VAR_OUTPUT
    bIndexReq        : BOOL;                            // 分度请求，单拍脉冲 [-] [Index request, single-scan pulse]
    nActiveStation   : INT;                             // 当前作业工位号 [1~工位数]，0 表示无效 [Active station number, 0 = invalid]
    bStationReady    : BOOL;                            // 当前工位允许工艺动作 [-] [Station ready for process action]
    nRecipeAtStation : INT;                             // 当前工位工艺号，透传 [-] [Recipe number at active station]
    uStationMask     : DWORD;                           // 工位启用镜像，第 n 位对应第 n 工位 [Station enable mirror, bit n-1]
    bCycleDone       : BOOL;                            // 整圈走完单拍脉冲 [-] [Single pulse on full revolution]
    tDwellRemain     : TIME;                            // 当前工位剩余停留时间 [毫秒] [Remaining dwell time]
    eState           : E_DL_IndexTableState;            // 主状态机当前态 [-] [Current state]
    bError           : BOOL;                            // 故障锁存，需复位清除 [Latched fault]
    uErrorId         : UDINT;                           // 事件码或故障码，0 表示无 [Event or fault code]
END_VAR
VAR_IN_OUT
    stStat           : ST_DL_IndexTableStat;            // 跨周期统计，调用方持有 [Persistent statistics]
END_VAR
VAR
    _eState          : E_DL_IndexTableState := E_DL_IndexTableState.eIdle;  // 内部状态寄存器，唯一真值源 [Internal state register]
    _bInit           : BOOL := FALSE;                   // 首扫标志，初值 FALSE，判据 NOT _bInit [First-scan flag, R19 pattern]
    _bFaultLatch     : BOOL;                            // 故障级锁存，仅复位路径清 [Fault latch, reset path only]
    _uErrorIdInt     : UDINT;                           // 故障级码寄存 [Fault-level code register]
    _uInfoCode       : UDINT;                           // 本拍信息级码，每拍重算 [Transient info code]
    nStaEff          : INT;                             // 生效工位数，已钳位 [个] [Effective station count]
    nIdxVal          : INT;                             // 到位工位号（已判界）[号] [Validated station number]
    tDwellEff        : TIME;                            // 生效停留时间 [毫秒] [Effective dwell time]
    tSettleEff       : TIME;                            // 生效稳定时间 [毫秒] [Effective settling time]
    tIndexEff        : TIME;                            // 生效分度超时 [毫秒] [Effective index timeout]
    tCycleEff        : TIME;                            // 生效扫描周期 [毫秒] [Effective task cycle time]
    uMaskAcc         : UDINT;                           // 掩码累加器 [位域] [Mask accumulator]
    uBitAcc          : UDINT;                           // 位累加器，逐位左移 [位域] [Single-bit accumulator]
    nI               : INT;                             // 通用循环索引 [索引] [Loop index]
    bDwellIn         : BOOL;                            // 停留计时输入条件，先算后调 [Dwell timer input]
    bSettleIn        : BOOL;                            // 稳定计时输入条件，先算后调 [Settle timer input]
    bIndexIn         : BOOL;                            // 分度超时输入条件，先算后调 [Index timer input]
    bDwellDone       : BOOL;                            // 停留结束（含空跑旁路）[Dwell finished, dry-run bypassed]
    _bInPosDropped   : BOOL;                            // 分度中到位信号曾回落，兼容保持型开关 [In-position dropped during indexing]
    fbTrigStart      : R_TRIG;                          // 启动沿检测 [Start edge detector]
    fbTrigStop       : R_TRIG;                          // 停止沿检测 [Stop edge detector]
    fbTrigReset      : R_TRIG;                          // 复位沿检测 [Reset edge detector]
    fbTrigInPos      : R_TRIG;                          // 到位上升沿检测 [In-position rising edge]
    fbTrigInPosFall  : F_TRIG;                          // 到位下降沿检测，抖动诊断用 [In-position falling edge, jitter diagnosis]
    fbTmoDwell       : TON;                             // 停留计时 [Dwell timer]
    fbTmoSettle      : TON;                             // 稳定确认计时 [Settle timer]
    fbTmoIndex       : TON;                             // 分度超时 [Index timeout timer]
END_VAR
VAR CONSTANT
    DL_STATION_MAX   : INT := 24;                       // 工位上限 [个] [Max station count]
    DL_STATION_MIN   : INT := 2;                        // 工位下限 [个] [Min station count]
    DL_TMO_MAX       : TIME := T#120S;                  // 时长参数域上限 [毫秒] [Duration upper bound]
    DL_RUN_MAX       : TIME := T#500H;                 // 运行时长饱和上限 [毫秒] [Run time saturation limit]
    DL_COUNT_MAX     : UDINT := 16#FFFF_FFFE;           // 计数饱和上限 [次] [Counter saturation limit]
    DL_INFO_STA_CLAMP: UDINT := 16#0005_01C2;           // 01C2 工位数量越界已钳位【信息级】 [Info, station count clamped]
    DL_ERR_INDEX_TMO : UDINT := 16#0005_02D0;           // 02D0 分度超时【故障级】 [Fault, index timeout]
    DL_ERR_INPOS     : UDINT := 16#0005_02D1;           // 02D1 到位信号抖动或丢失【故障级】 [Fault, in-position lost]
    DL_ERR_STATION   : UDINT := 16#0005_02D2;           // 02D2 工位号越界【故障级】 [Fault, station out of range]
    DL_ERR_STATE     : UDINT := 16#0005_02D3;           // 02D3 非法状态兜底【故障级】 [Fault, illegal state]
END_VAR

// ==== 段 1｜单拍输出预清零（脉冲类出口每拍先清零，避免跨拍粘滞） / Single-scan pulse pre-clear, no sticky pulses
bIndexReq  := FALSE;                        // 分度请求先清零 [Index request pre-cleared]
bCycleDone := FALSE;                        // 整圈完成先清零 [Revolution pulse pre-cleared]
_uInfoCode := 16#0000_0000;                 // 信息级码每拍重算 [Info code recomputed]

// ==== 段 2｜参数钳位（工位数与三个时长，先钳位再进逻辑） / Parameter clamping before any logical use
nStaEff := nStationCount;                   // 工位数先取引脚值 [Station count from pin]
IF nStaEff < DL_STATION_MIN THEN
    nStaEff    := DL_STATION_MIN;           // 低于下限钳到 2 [Clamped to lower bound]
    _uInfoCode := DL_INFO_STA_CLAMP;        // 01C2 工位数量越界已钳位【信息级】 [Info, count clamped]
ELSIF nStaEff > DL_STATION_MAX THEN
    nStaEff    := DL_STATION_MAX;           // 高于上限钳到 24 [Clamped to upper bound]
    _uInfoCode := DL_INFO_STA_CLAMP;        // 01C2 工位数量越界已钳位【信息级】 [Info, count clamped]
END_IF

tDwellEff := tDwellTime;                    // 停留时间先取引脚值 [Dwell from pin]
IF tDwellEff > DL_TMO_MAX THEN
    tDwellEff := DL_TMO_MAX;                // 超上限钳位 [Clamped to upper bound]
ELSIF tDwellEff < T#0S THEN
    tDwellEff := T#0S;                      // 负值归零 [Negative clamped to zero]
END_IF

tSettleEff := tSettleTime;                  // 稳定时间先取引脚值 [Settle from pin]
IF tSettleEff > DL_TMO_MAX THEN
    tSettleEff := DL_TMO_MAX;               // 超上限钳位 [Clamped to upper bound]
ELSIF tSettleEff < T#0S THEN
    tSettleEff := T#0S;                     // 负值归零 [Negative clamped to zero]
END_IF

tIndexEff := tIndexTimeout;                 // 分度超时先取引脚值 [Index timeout from pin]
IF tIndexEff > DL_TMO_MAX THEN
    tIndexEff := DL_TMO_MAX;                // 超上限钳位 [Clamped to upper bound]
ELSIF tIndexEff <= T#0S THEN
    tIndexEff := T#0S;                      // 零表示不监控 [Zero means supervision disabled]
END_IF

tCycleEff := tCycle;                        // 扫描周期先取引脚值 [Task cycle from pin]
IF tCycleEff <= T#0S OR tCycleEff > T#10S THEN
    tCycleEff := T#10MS;                    // 异常值回默认 10 毫秒 [Fallback to 10 ms]
END_IF

// ==== 段 3｜沿与定时器无条件刷新（R7 红线：严禁置于 IF / CASE 分支内） / Unconditional refresh of edges and timers
fbTrigStart(CLK := bStart);                 // 启动沿 [Start edge]
fbTrigStop(CLK := bStop);                   // 停止沿 [Stop edge]
fbTrigReset(CLK := bReset);                 // 复位沿 [Reset edge]
fbTrigInPos(CLK := bIndexInPos);            // 到位上升沿 [In-position rising edge]
fbTrigInPosFall(CLK := bIndexInPos);        // 到位下降沿 [In-position falling edge]

IF _eState = E_DL_IndexTableState.eDwell THEN
    bDwellIn := TRUE;                       // 仅停留段计时 [Only during dwell]
ELSE
    bDwellIn := FALSE;                      // 其余段清零 [Cleared otherwise]
END_IF
fbTmoDwell(IN := bDwellIn, PT := tDwellEff);

IF _eState = E_DL_IndexTableState.eSettling THEN
    bSettleIn := TRUE;                      // 仅稳定段计时 [Only during settling]
ELSE
    bSettleIn := FALSE;                     // 其余段清零 [Cleared otherwise]
END_IF
fbTmoSettle(IN := bSettleIn, PT := tSettleEff);

IF (_eState = E_DL_IndexTableState.eIndexing) AND (tIndexEff > T#0S) THEN
    bIndexIn := TRUE;                       // 仅分度段且监控开启时计时 [Only while indexing with supervision on]
ELSE
    bIndexIn := FALSE;                      // 其余段清零 [Cleared otherwise]
END_IF
fbTmoIndex(IN := bIndexIn, PT := tIndexEff);

// ==== 段 4｜首扫初始化（R19 唯一合法范式：初值 FALSE，判据 NOT，同步后置 TRUE） / First-scan initialisation with the canonical R19 pattern
IF NOT _bInit THEN
    _eState          := E_DL_IndexTableState.eIdle;  // 状态回待机 [State to idle]
    _bInPosDropped   := FALSE;              // 到位回落标志复位 [Dropped flag reset]
    _bFaultLatch     := FALSE;              // 故障锁存清零 [Fault latch cleared]
    _uErrorIdInt     := 16#0000_0000;       // 故障码清零 [Fault code cleared]
    nActiveStation   := 0;                  // 作业工位号清 0 [Active station cleared]
    nRecipeAtStation := 0;                  // 工艺号清 0 [Recipe cleared]
    bStationReady    := FALSE;              // 放行复位 [Permit cleared]
    tDwellRemain     := T#0S;               // 剩余停留清零 [Remaining dwell cleared]
    bError           := FALSE;              // 故障标志清零 [Error cleared]
    uErrorId         := 16#0000_0000;       // 事件码清零 [Error id cleared]
    stStat.nIndexCount := 0;                // 分度计数清零 [Index counter cleared]
    stStat.nCycleCount := 0;                // 循环计数清零 [Revolution counter cleared]
    stStat.tRunTime    := T#0S;             // 运行时长清零 [Run time cleared]
    _bInit := TRUE;                         // 首扫只做一次 [Runs exactly once]
END_IF

// ==== 段 5｜工位启用掩码重建（逐位置位，不用累计量拼接，规避位宽边界） / Mask rebuild by per-bit set, no shift accumulation
uMaskAcc := 0;
uBitAcc  := 1;
FOR nI := 1 TO DL_STATION_MAX DO
    IF (nI <= nStaEff) AND abStationEnable[nI] THEN
        uMaskAcc := uMaskAcc OR uBitAcc;    // 该工位启用则置对应位 [Set bit for enabled station]
    END_IF
    uBitAcc := uBitAcc * 2;                 // 位累加器左移一位（等价左移，跨平台不依赖位移函数）[Shift left by one]
END_FOR
uStationMask := UDINT_TO_DWORD(uMaskAcc);   // 转位串出口 [Convert to word for output]

// ==== 段 6｜使能撤销（FALSE 立即回待机、撤分度请求、清作业工位） / Disable path withdraws the request and clears the station
IF NOT bEnable THEN
    _eState        := E_DL_IndexTableState.eIdle;
    bIndexReq      := FALSE;                // 请求撤销 [Request withdrawn]
    bStationReady  := FALSE;                // 放行撤销 [Permit withdrawn]
    nActiveStation := 0;                    // 作业工位清 0 [Active station cleared]
END_IF

// ==== 段 7｜全局监视：工位号越界在分度链之外单点判定，避免越界索引数组 / Bounds monitor outside the CASE, protects array access
IF bEnable AND (NOT _bFaultLatch)
AND (_eState <> E_DL_IndexTableState.eIdle)
AND (_eState <> E_DL_IndexTableState.eFault)
AND ((nAtStation < 0) OR (nAtStation > nStaEff)) THEN
    bIndexReq    := FALSE;                  // 越界即撤请求 [Request withdrawn on out-of-range]
    _bFaultLatch := TRUE;                   // 故障锁存 [Fault latched]
    _uErrorIdInt := DL_ERR_STATION;         // 02D2 工位号越界【故障级】 [Fault, station out of range]
    _eState      := E_DL_IndexTableState.eFault;
END_IF

// ==== 段 8｜主状态机（ENUM 加 CASE 加 ELSE 兜底，五成员逐一有标签） / Main state machine, every member has its own label
CASE _eState OF
    E_DL_IndexTableState.eIdle: // 待机：等启动沿，首工位放行由停留态给出
        IF fbTrigStart.Q AND bEnable AND (NOT _bFaultLatch) THEN
            _uErrorIdInt := 16#0000_0000;   // 启动前必无故障，码清零 [No fault before start]
            IF (nAtStation >= 1) AND (nAtStation <= nStaEff) THEN
                nActiveStation := nAtStation;   // 已定位则先放行该工位 [Permit current station if seated]
            ELSE
                nActiveStation := 0;        // 未定位不给放行 [No permit when not seated]
            END_IF
            _eState := E_DL_IndexTableState.eDwell;
        END_IF

    E_DL_IndexTableState.eDwell: // 停留：工艺放行窗，计时到即出分度请求
        IF (nAtStation >= 1) AND (nAtStation <= nStaEff) THEN
            nActiveStation := nAtStation;       // 作业工位跟随机械反馈 [Follow mechanical feedback]
        ELSE
            nActiveStation := 0;                // 未定位则无效 [Invalid when not seated]
        END_IF
        IF bDryRun THEN
            bDwellDone := TRUE;                 // 空跑旁路停留计时 [Dry run bypasses dwell]
        ELSE
            bDwellDone := fbTmoDwell.Q;         // 正常按定时器 [Normal timer]
        END_IF
        IF bDwellDone THEN
            IF fbTrigStop.Q OR bStop THEN    // 上升沿受理短脉冲按钮，电平兜住长按与上位机置位 [Edge for momentary, level for held stop]
                _eState := E_DL_IndexTableState.eIdle;   // 停止请求：完成当前工位后停 [Stop after current station]
            ELSE
                bIndexReq      := TRUE;         // 分度请求单拍脉冲，本拍唯一置位点 [Sole set point of the pulse]
                _bInPosDropped := FALSE;        // 新的分度周期，回落标志复位 [Dropped flag reset per index]
                _eState        := E_DL_IndexTableState.eIndexing;
            END_IF
        END_IF

    E_DL_IndexTableState.eIndexing: // 分度中：等到位确认，超时即锁故障
        IF NOT bIndexInPos THEN
            _bInPosDropped := TRUE;             // 到位信号已回落，后续恢复即可确认 [Signal dropped, recovery confirms]
        END_IF
        IF fbTrigInPos.Q OR (_bInPosDropped AND bIndexInPos) THEN
            IF stStat.nIndexCount < DL_COUNT_MAX THEN
                stStat.nIndexCount := stStat.nIndexCount + 1;  // 成功分度计数（偏离 D2）[Successful index counter]
            END_IF
            _eState := E_DL_IndexTableState.eSettling;
        ELSIF fbTmoIndex.Q THEN
            _bFaultLatch := TRUE;               // 超时锁存 [Timeout latched]
            _uErrorIdInt := DL_ERR_INDEX_TMO;   // 02D0 分度超时【故障级】 [Fault, index timeout]
            _eState      := E_DL_IndexTableState.eFault;
        END_IF

    E_DL_IndexTableState.eSettling: // 稳定中：去抖确认，掉沿即判硬件抖动
        IF fbTrigInPosFall.Q THEN
            _bFaultLatch := TRUE;               // 抖动属硬件问题，锁故障且不重试 [Hardware fault, no retry]
            _uErrorIdInt := DL_ERR_INPOS;       // 02D1 到位信号抖动或丢失【故障级】 [Fault, in-position lost]
            _eState      := E_DL_IndexTableState.eFault;
        ELSIF (nAtStation < 1) OR (nAtStation > nStaEff) THEN
            _bFaultLatch := TRUE;               // 稳定窗内工位号失真 [Station feedback untrustworthy]
            _uErrorIdInt := DL_ERR_STATION;     // 02D2 工位号越界【故障级】 [Fault, station out of range]
            _eState      := E_DL_IndexTableState.eFault;
        ELSIF bIndexInPos AND fbTmoSettle.Q THEN
            nActiveStation := nAtStation;       // 稳定通过，登记作业工位 [Settled, register active station]
            IF (NOT bDryRun) AND (nAtStation = 1) THEN
                bCycleDone := TRUE;             // 回到 1 号位即整圈完成单拍 [Sole set point of the pulse]
                IF stStat.nCycleCount < DL_COUNT_MAX THEN
                    stStat.nCycleCount := stStat.nCycleCount + 1;  // 循环计数饱和累加 [Revolution counter, saturated]
                END_IF
            END_IF
            _eState := E_DL_IndexTableState.eDwell;
        END_IF

    E_DL_IndexTableState.eFault: // 故障：等复位沿，复位后清码回待机
        bIndexReq      := FALSE;                // 故障态不得出请求 [No request while faulted]
        bStationReady  := FALSE;                // 故障态不得放行 [No permit while faulted]
        IF fbTrigReset.Q THEN
            _bFaultLatch   := FALSE;            // 锁存解除 [Latch released]
            _bInPosDropped := FALSE;            // 到位回落标志复位 [Dropped flag reset]
            _uErrorIdInt   := 16#0000_0000;     // 故障码清零 [Fault code cleared]
            nActiveStation := 0;                // 作业工位清 0 [Active station cleared]
            _eState      := E_DL_IndexTableState.eIdle;
        END_IF

    ELSE // 非法枚举值兜底：撤请求、回安全态并锁故障
        bIndexReq    := FALSE;                  // 非法态撤请求 [Request withdrawn]
        _bFaultLatch := TRUE;                   // 兜底锁存 [Fallback latch]
        _uErrorIdInt := DL_ERR_STATE;           // 02D3 非法状态兜底【故障级】 [Fault, illegal state]
        _eState      := E_DL_IndexTableState.eFault;
END_CASE

// ==== 段 9｜运行时长累计（仅运行段累加，饱和保护，停机不计） / Run-time accumulation with saturation
IF bEnable AND (_eState <> E_DL_IndexTableState.eIdle)
AND (_eState <> E_DL_IndexTableState.eFault)
AND (stStat.tRunTime < DL_RUN_MAX) THEN
    stStat.tRunTime := stStat.tRunTime + tCycleEff;   // 累加一个扫描周期 [Accumulate one task cycle]
END_IF

// ==== 段 10｜出口派生（放行、工艺号、剩余停留三者在同一处单点派生） / Outlets derived at a single point
bStationReady := FALSE;                    // 默认不放行，判界通过后再置位 [Default no permit, bounds checked first]
IF (NOT bDryRun) AND (_eState = E_DL_IndexTableState.eDwell)
AND (nActiveStation >= 1) AND (nActiveStation <= nStaEff) THEN
    bStationReady := abStationEnable[nActiveStation];   // 放行：工位启用才放 [Permit only when the station is enabled]
END_IF

IF (nActiveStation >= 1) AND (nActiveStation <= nStaEff) THEN
    nRecipeAtStation := anStationRecipe[nActiveStation];   // 工艺号透传 [Recipe pass-through]
ELSE
    nRecipeAtStation := 0;                  // 无效工位给 0 [Zero for invalid station]
END_IF

IF tDwellEff > fbTmoDwell.ET THEN
    tDwellRemain := tDwellEff - fbTmoDwell.ET;   // 剩余停留时间 [Remaining dwell]
ELSE
    tDwellRemain := T#0S;                   // 已到点钳零 [Clamped to zero]
END_IF

eState  := _eState;                         // 状态镜像 [State mirror]
bError  := _bFaultLatch;                    // 故障级派生式（R21）[Fault-level derived form]
IF _bFaultLatch THEN
    uErrorId := _uErrorIdInt;               // 故障级码优先透出 [Fault code wins]
ELSE
    uErrorId := _uInfoCode;                 // 无故障时透出信息级码 [Info code otherwise]
END_IF
END_FUNCTION_BLOCK

(* ---- FB_DL_SlurryMixingSeq.st ---- *)
(*==============================================================================
 * 组件名称 (Component)  : FB_DL_SlurryMixingSeq
 * 所属子库 (Sublibrary) : DL_Process
 * 当前版本 (Version)    : 1.0.0
 * 兼容性   (Platform)   : CODESYS 3.5+ / TwinCAT 3 / 汇川 InoProShop / 施耐德 Machine Expert
 *                         仅依赖 Standard.library（TON / R_TRIG / ABS），零厂商私有库
 * 功能描述 (Function)   : 浆料批次四相顺控：eIdle → eFill（加料，料位或重量达窗）→ eDisperse
 *                         （高速分散：转速达窗 + 分散时长 tDisperse）→ eDeair（真空脱泡：真空度
 *                         达窗 + 脱泡时长 tDeair）→ eDischarge（出料：料位到下限或撤启动）→ eDone。
 *                         相内监视：温升速率超 fTempRiseMax 立即故障（浆料过热会凝胶，属安全侧
 *                         异常，按 R146 立即终止）；分散相时长届满时转速仍在容差带外 → 失速故障。
 *                         每相独立超时（tFillMax / tDisperseMax / tDeairMax / tDischargeMax）。
 * 撤启动语义 (Abort)    : **bStart 落沿在任意执行相 → 直接进 eDischarge 安全收料**，不得停在
 *                         分散相（分散中滞留会让浆料在高速剪切下持续升温）。这是 R98 双出口
 *                         范式在本件的落地：执行相均有「工艺达成」与「撤启动」两条出口。
 * 分工声明 (Scope)      : 与 `FB_DL_SlurryStirrerCtrl`（Device 子库，单机搅拌器驱动与转速
 *                         闭环）分工 —— 本件是**批次相序编排**，只发相级命令位，不直接驱动
 *                         电机、不做转速闭环。
 * 接口     (Interface)  : 输入 bStart 启动电平、料位/重量/转速/真空/温升与各自目标与容差、
 *                         四个工艺时长与四个相超时、bReset 复位；输出 eState 相位、eCause 归因、
 *                         四个相级命令位、bCycleDone 完成标志、bError / nErrId。
 * 边界     (Boundary)   : ① 组态闸：任一容差 <= 0.0、任一时长 <= T#0S、fLevelHiPct <= fLevelLoPct、
 *                         fWeightTgtKg <= 0.0、fVacTgtKpa <= 0.0、fTempRiseMax <= 0.0 或任一浮点
 *                         引脚 NaN → 故障锁存（每个参与判据的引脚都在闸内，R151）；
 *                         ② **4 枚 TON（相计时）+ 1 枚 R_TRIG 全部段 0 无条件刷新**，每个实例的
 *                         IN 由对应相位派生（R228A），离开该相 IN 落假 → Q 落假、ET 归零
 *                         （R228B 跨相复位语义成立）；本件是本轮 TON 密度最高件，逐实例已核：
 *                         tonFill↔eFill、tonDisperse↔eDisperse、tonDeair↔eDeair、
 *                         tonDischarge↔eDischarge，四者对相位一一绑定，无跨相复用；
 *                         ③ 相时长的「工艺时间」与「相超时」共用同一实例：PT 绑该相超时上限，
 *                         工艺达成判据读 ET（ET >= 工艺时长），结构上不可能出现「两个计时器
 *                         各说各话」；④ 故障相迁出唯一路径 = bReset 上升沿；
 *                         ⑤ 零全局耦合（无 GVL / 无物理地址）。
 * 解除式   (Release)    : bReset 上升沿 ∧ 组态合法 ∧ 已撤启动（NOT bStart，当拍量，R240 范式）。
 *                         自证可满足（终审两式 1）：四枚 TON 的 IN 挂相位，故障相内 IN 恒假 →
 *                         Q 恒假；bStart 为外部电平，操作员松开即达，无恒假因子。
 * 码表     (Codes)      : 16#0005_03A6 故障级：浆料混合顺控故障总码（组态非法 / 加料超时 /
 *                         转速失速 / 真空不足 / 温升超限 / 出料超时 / 非法相位），锁存至 bReset
 *                         上升沿，归因由 eCause 承载（R190 单件单总码，每个成因均有独立赋值点）；
 *                         16#0005_04CE 信息级：批次循环完成（进 eDone 单拍）。
 *                         加码反证（R90）：完成时 bCycleDone 由相位派生且四命令位全落，而「长时间
 *                         停在 eDone」与之同值，出口组合无法区分「刚完成一个批次」与「完成态驻留」，
 *                         故立一码记录每个批次的完成沿。
 *                         码段说明：0005 段故障子带 03xx / 信息子带 04xx，本件取 03A6 / 04CE
 *                         （源码实扫该两槽为空，续接同子带已用最大值，未回填碎片孔洞）。
 * 开源溯源 (Origin)     : 道莅自研 clean-room（参考锂电前段浆料制备工艺与公开参数域，
 *                         零代码行复制；自研行业池）
 * 修订历史 (Revision)   : 2026-11-19  v1.0.0  R45 首版（批次 4 · 序号 18）
 *==============================================================================*)

TYPE E_DL_SmxState :
(
    eIdle      := 0,     // 待启动 / Idle, awaiting start
    eFill      := 10,    // 加料相 / Filling
    eDisperse  := 20,    // 高速分散相 / High-speed dispersion
    eDeair     := 30,    // 真空脱泡相 / Vacuum de-airing
    eDischarge := 40,    // 出料相（含撤启动安全收料） / Discharging, also the safe abort target
    eDone      := 50,    // 批次完成 / Batch done
    eFault     := 90     // 故障锁存相 / Fault latched phase
);
END_TYPE

TYPE E_DL_SmxCause :
(
    eNone         := 0,  // 无故障成因 / No cause
    eCfgIllegal   := 1,  // 组态非法 / Illegal configuration
    eFillTmo      := 2,  // 加料超时 / Fill timeout
    eSpeedLoss    := 3,  // 转速失速（时长届满仍在容差带外） / Speed out of tolerance at time-up
    eVacLow       := 4,  // 真空不足 / Vacuum insufficient
    eTempRise     := 5,  // 温升速率超限 / Temperature rise rate over limit
    eDischargeTmo := 6,  // 出料超时 / Discharge timeout
    ePhaseBad     := 7   // 非法相位兜底 / Illegal phase fallback
);
END_TYPE

FUNCTION_BLOCK FB_DL_SlurryMixingSeq
VAR_INPUT
    bStart        : BOOL := FALSE;        // 批次启动电平（落沿触发安全收料） [-] / Batch start level, falling edge triggers safe discharge
    fLevelPct     : REAL := 0.0;          // 料位 [%] / Tank level [%]
    fLevelLoPct   : REAL := 5.0;          // 料位下限（出料终点），域 < fLevelHiPct [%] / Level low limit [%]
    fLevelHiPct   : REAL := 80.0;         // 料位上限（加料终点），域 > fLevelLoPct [%] / Level high limit [%]
    fWeightKg     : REAL := 0.0;          // 批次重量 [kg] / Batch weight [kg]
    fWeightTgtKg  : REAL := 500.0;        // 目标重量，域 > 0.0 [kg] / Target weight, domain > 0.0 [kg]
    fSpeedRpm     : REAL := 0.0;          // 实测转速 [rpm] / Measured speed [rpm]
    fSpeedTgtRpm  : REAL := 1200.0;       // 分散目标转速 [rpm] / Dispersion target speed [rpm]
    fSpeedTol     : REAL := 50.0;         // 转速容差带，域 > 0.0 [rpm] / Speed tolerance, domain > 0.0 [rpm]
    fVacKpa       : REAL := 0.0;          // 实测真空度（幅值） [kPa] / Measured vacuum magnitude [kPa]
    fVacTgtKpa    : REAL := 80.0;         // 真空目标（幅值），域 > 0.0 [kPa] / Vacuum target magnitude, domain > 0.0 [kPa]
    fTempRiseCpm  : REAL := 0.0;          // 温升速率 [°C/min] / Temperature rise rate [degC/min]
    fTempRiseMax  : REAL := 2.0;          // 温升速率上限，域 > 0.0 [°C/min] / Rise-rate limit, domain > 0.0 [degC/min]
    tFill         : TIME := T#30S;        // 加料最短时长（防料位抖动误判），域 > T#0S [ms] / Fill minimum duration [ms]
    tFillMax      : TIME := T#10M;        // 加料相超时，域 > tFill [ms] / Fill phase timeout [ms]
    tDisperse     : TIME := T#20M;        // 分散工艺时长，域 > T#0S [ms] / Dispersion process time [ms]
    tDisperseMax  : TIME := T#25M;        // 分散相超时，域 > tDisperse [ms] / Dispersion phase timeout [ms]
    tDeair        : TIME := T#15M;        // 脱泡工艺时长，域 > T#0S [ms] / De-airing process time [ms]
    tDeairMax     : TIME := T#20M;        // 脱泡相超时，域 > tDeair [ms] / De-airing phase timeout [ms]
    tDischarge    : TIME := T#30S;        // 出料最短时长，域 > T#0S [ms] / Discharge minimum duration [ms]
    tDischargeMax : TIME := T#5M;         // 出料相超时，域 > tDischarge [ms] / Discharge phase timeout [ms]
    bReset        : BOOL := FALSE;        // 复位命令，上升沿清故障 [-] / Reset command, rising edge clears fault
END_VAR
VAR_OUTPUT
    eState            : E_DL_SmxState;    // 状态出口，段 6 单点映射 / State outlet
    eCause            : E_DL_SmxCause;    // 故障成因出口（R190 归因唯一） / Fault cause outlet
    bInletValveCmd    : BOOL;             // 进料阀命令（仅加料相） [-] / Inlet valve command, fill phase only
    bStirrerFastCmd   : BOOL;             // 高速搅拌命令（分散相） [-] / High-speed stirrer command, disperse phase
    bVacPumpCmd       : BOOL;             // 真空泵命令（脱泡相） [-] / Vacuum pump command, de-air phase
    bDischargeValveCmd: BOOL;             // 出料阀命令（出料相） [-] / Discharge valve command, discharge phase
    bCycleDone        : BOOL;             // 批次完成标志 [-] / Batch done flag
    bError            : BOOL;             // 故障锁存标志 [-] / Fault latch flag
    nErrId            : UDINT;            // 事件码，0 = 无事件 / Event code, 0 = no event
END_VAR
VAR
    _eState       : E_DL_SmxState := E_DL_SmxState.eIdle;   // 内部相位（CASE 唯一写入目标） / Internal phase
    _eCause       : E_DL_SmxCause := E_DL_SmxCause.eNone;   // 故障成因锁存（锁存量） / Latched cause
    tonFill       : TON;                  // 加料相计时（PT = 相超时），段 0 无条件调用 / Fill phase timer
    tonDisperse   : TON;                  // 分散相计时（PT = 相超时），段 0 无条件调用 / Dispersion phase timer
    tonDeair      : TON;                  // 脱泡相计时（PT = 相超时），段 0 无条件调用 / De-air phase timer
    tonDischarge  : TON;                  // 出料相计时（PT = 相超时），段 0 无条件调用 / Discharge phase timer
    rtReset       : R_TRIG;               // 复位沿实例，段 0 无条件调用 / Reset edge
    _bSpeedInTol  : BOOL;                 // 转速在容差带当拍量 [-] / Speed inside tolerance
    _bVacInTol    : BOOL;                 // 真空达窗当拍量 [-] / Vacuum reached
    _bFillReached : BOOL;                 // 加料达窗当拍量 [-] / Fill reached
    _bDischDone   : BOOL;                 // 出料完成当拍量 [-] / Discharge finished
    _bNonFin      : BOOL;                 // 输入非有限当拍量 [-] / Non-finite input this scan
    _bCfgBad      : BOOL;                 // 组态非法当拍量 [-] / Illegal configuration
    _bFault       : BOOL;                 // 故障锁存位（锁存量） / Latched fault bit
    _uFault       : UDINT;                // 故障码锁存（锁存量） / Latched fault code
    _uInfo        : UDINT;                // 信息码，每拍重算 / Info code, recomputed each scan
END_VAR
VAR CONSTANT
    DL_SPEED_EPS : REAL := 1.0E-3;        // 判据辅助容差（防阈值给出极小值时的边界抖动） [无量纲] / Criterion epsilon [dimensionless]
END_VAR

(* —— 段 0：当拍判据派生 + 4 枚 TON 与沿实例无条件周期刷新（逐实例绑定相位） —— *)
_bNonFin := (fLevelPct <> fLevelPct) OR (fWeightKg <> fWeightKg) OR (fSpeedRpm <> fSpeedRpm)      // NaN 自反判（判等禁令唯一例外） / NaN self-reflexive tests
         OR (fVacKpa <> fVacKpa) OR (fTempRiseCpm <> fTempRiseCpm);                                // 真空与温升 NaN 判 / Vacuum and rise-rate NaN tests
_bSpeedInTol  := ABS(fSpeedRpm - fSpeedTgtRpm) <= (fSpeedTol + DL_SPEED_EPS);                      // 转速容差判据 / Speed tolerance verdict
_bVacInTol    := fVacKpa >= (fVacTgtKpa - DL_SPEED_EPS);                                            // 真空达窗判据 / Vacuum reached verdict
_bFillReached := (fLevelPct >= (fLevelHiPct - DL_SPEED_EPS)) OR (fWeightKg >= (fWeightTgtKg - DL_SPEED_EPS));   // 料位或重量达窗 / Level or weight reached
_bDischDone   := fLevelPct <= (fLevelLoPct + DL_SPEED_EPS);                                         // 料位到下限 / Level reached low limit
_bCfgBad := (fSpeedTol <= 0.0) OR (fTempRiseMax <= 0.0) OR (fLevelHiPct <= fLevelLoPct)             // 容差与料位几何闸 / Tolerance and level geometry gates
            OR (fWeightTgtKg <= 0.0) OR (fVacTgtKpa <= 0.0)                                         // 重量与真空目标正域闸 / Weight and vacuum gates
            OR (tFill <= T#0S) OR (tFillMax <= tFill) OR (tDisperse <= T#0S) OR (tDisperseMax <= tDisperse)   // 时间正域与配比闸 / Time gates and ratio constraints
            OR (tDeair <= T#0S) OR (tDeairMax <= tDeair)                                            // 脱泡时间配比闸 / De-air time gates
            OR (tDischarge <= T#0S) OR (tDischargeMax <= tDischarge);                               // 出料时间配比闸 / Discharge time gates
rtReset(CLK := bReset);                                                                             // 复位沿，每拍必调（R228A） / Reset edge
tonFill(IN := (_eState = E_DL_SmxState.eFill), PT := tFillMax);                                     // 加料相计时（IN 绑相位） / Fill timer, phase-bound
tonDisperse(IN := (_eState = E_DL_SmxState.eDisperse), PT := tDisperseMax);                         // 分散相计时（IN 绑相位） / Dispersion timer, phase-bound
tonDeair(IN := (_eState = E_DL_SmxState.eDeair), PT := tDeairMax);                                  // 脱泡相计时（IN 绑相位） / De-air timer, phase-bound
tonDischarge(IN := (_eState = E_DL_SmxState.eDischarge), PT := tDischargeMax);                      // 出料相计时（IN 绑相位） / Discharge timer, phase-bound

(* —— 段 1：单拍量预清零（锁存量不入清单，R107） —— *)
_uInfo   := 16#0000_0000;          // 信息码每拍重算 / Info recomputed every scan
nErrId   := 16#0000_0000;          // 事件码缺省无事件 / Event code default none
bError   := FALSE;                 // 故障标志每拍预清，故障分支同拍置位（R45 配对） / Flag preset

(* —— 段 2：复位沿 + 组态域闸 + 非有限闸 —— *)
IF rtReset.Q THEN                                                        // 当拍复位沿 / current-scan reset edge
    _bFault := FALSE;                                                    // 清故障锁存位（锁存量） / Clear fault latch
    _uFault := 16#0000_0000;                                             // 清故障锁存码（锁存量） / Clear latched code
    _eCause := E_DL_SmxCause.eNone;                                      // 清成因（锁存量） / Clear latched cause
    IF _eState = E_DL_SmxState.eFault THEN
        _eState := E_DL_SmxState.eIdle;                                  // 故障相迁出唯一路径 / Sole exit from fault phase
    END_IF
END_IF
IF _bCfgBad THEN                                                         // 组态域闸 / Configuration gate
    _uFault := 16#0005_03A6;                                             // 故障级：浆料混合顺控故障总码 / Fault-level: slurry sequence fault code
    _bFault := TRUE;
    bError  := TRUE;                                                     // 故障标志同拍置位（R45 配对） / Error flag set same scan
    _eCause := E_DL_SmxCause.eCfgIllegal;                                // 归因：组态非法 / Cause: illegal configuration
END_IF
IF (NOT _bFault) AND _bNonFin THEN                                       // 输入非有限（归入组态非法归因） / Non-finite input, mapped to config cause
    _uFault := 16#0005_03A6;
    _bFault := TRUE;
    bError  := TRUE;
    _eCause := E_DL_SmxCause.eCfgIllegal;                                // 归因：组态非法（含非有限输入） / Cause: illegal configuration including non-finite
END_IF

(* —— 段 3：温升速率监视（安全侧异常，立即终止，R146） —— *)
IF (NOT _bFault) AND (fTempRiseCpm > fTempRiseMax) THEN
    _uFault := 16#0005_03A6;                                             // 故障级：温升超限 / Fault-level: rise rate over limit
    _bFault := TRUE;
    bError  := TRUE;
    _eCause := E_DL_SmxCause.eTempRise;                                  // 归因：温升超限 / Cause: temperature rise
END_IF

(* —— 段 4：相超时与相内判据（各成因独立赋值点，R190） —— *)
IF (NOT _bFault) AND tonFill.Q THEN                                      // 加料超时 / Fill timeout
    _uFault := 16#0005_03A6;
    _bFault := TRUE;
    bError  := TRUE;
    _eCause := E_DL_SmxCause.eFillTmo;                                   // 归因：加料超时 / Cause: fill timeout
END_IF
IF (NOT _bFault) AND tonDisperse.Q THEN                                  // 分散相时长届满仍失速 / Dispersion time-up with speed out of tolerance
    _uFault := 16#0005_03A6;
    _bFault := TRUE;
    bError  := TRUE;
    _eCause := E_DL_SmxCause.eSpeedLoss;                                 // 归因：转速失速 / Cause: speed loss
END_IF
IF (NOT _bFault) AND tonDeair.Q THEN                                     // 脱泡相时长届满真空仍不足 / De-air time-up with vacuum short
    _uFault := 16#0005_03A6;
    _bFault := TRUE;
    bError  := TRUE;
    _eCause := E_DL_SmxCause.eVacLow;                                    // 归因：真空不足 / Cause: vacuum insufficient
END_IF
IF (NOT _bFault) AND tonDischarge.Q THEN                                 // 出料超时 / Discharge timeout
    _uFault := 16#0005_03A6;
    _bFault := TRUE;
    bError  := TRUE;
    _eCause := E_DL_SmxCause.eDischargeTmo;                              // 归因：出料超时 / Cause: discharge timeout
END_IF

(* —— 段 5：故障解除式（R240 全当拍量） —— *)
IF rtReset.Q AND (NOT _bCfgBad) AND (NOT _bNonFin) AND (NOT bStart) THEN
    _bFault := FALSE;                                                    // 清故障锁存位（锁存量） / Clear fault latch
    _uFault := 16#0000_0000;                                             // 清故障锁存码（锁存量） / Clear latched code
    _eCause := E_DL_SmxCause.eNone;                                      // 清成因（锁存量） / Clear latched cause
END_IF

(* —— 段 5A：故障锁存相位迁移闸 —— *)
IF _bFault AND (_eState <> E_DL_SmxState.eFault) THEN
    _eState := E_DL_SmxState.eFault;                                     // 锁存即入故障相 / Latch enters fault phase
END_IF

(* —— 段 6：相位机（ENUM 全成员显式标签 + ELSE 兜底，R128） —— *)
CASE _eState OF

E_DL_SmxState.eIdle:
    IF bStart AND (NOT _bFault) THEN                                     // 出口 1：启动 / Start
        _eState := E_DL_SmxState.eFill;
    ELSIF _bFault THEN                                                   // 出口 2：故障锁存 / Fault latched
        _eState := E_DL_SmxState.eFault;
    END_IF

E_DL_SmxState.eFill:
    IF NOT bStart THEN                                                   // 出口 1：撤启动 → 安全收料（R98 双出口） / Start released, safe discharge
        _eState := E_DL_SmxState.eDischarge;
    ELSIF _bFillReached AND (tonFill.ET >= tFill) THEN                   // 出口 2：达窗且过最短时长 / Reached after minimum duration
        _eState := E_DL_SmxState.eDisperse;
    END_IF

E_DL_SmxState.eDisperse:
    IF NOT bStart THEN                                                   // 出口 1：撤启动 → 安全收料（R98 双出口） / Start released, safe discharge
        _eState := E_DL_SmxState.eDischarge;
    ELSIF _bSpeedInTol AND (tonDisperse.ET >= tDisperse) THEN            // 出口 2：转速达窗且分散时长满 / Speed reached and dispersion time done
        _eState := E_DL_SmxState.eDeair;
    END_IF

E_DL_SmxState.eDeair:
    IF NOT bStart THEN                                                   // 出口 1：撤启动 → 安全收料（R98 双出口） / Start released, safe discharge
        _eState := E_DL_SmxState.eDischarge;
    ELSIF _bVacInTol AND (tonDeair.ET >= tDeair) THEN                    // 出口 2：真空达窗且脱泡时长满 / Vacuum reached and de-air time done
        _eState := E_DL_SmxState.eDischarge;
    END_IF

E_DL_SmxState.eDischarge:
    IF _bDischDone AND (tonDischarge.ET >= tDischarge) THEN              // 出口 1：料位到下限且过最短时长 / Level low and minimum duration done
        _uInfo := 16#0005_04CE;                                          // 信息级：批次循环完成 / Info: batch completed
        _eState := E_DL_SmxState.eDone;
    ELSIF bStart THEN                                                    // 出口 2：重新给启动（前置消失，R98） / Start re-asserted
        _eState := E_DL_SmxState.eFill;
    END_IF

E_DL_SmxState.eDone:
    bCycleDone := TRUE;                                                  // 完成相保持完成标志 / Hold done flag in done phase
    IF NOT bStart THEN                                                   // 出口 1：撤启动回空闲 / Start released returns idle
        _eState := E_DL_SmxState.eIdle;
    ELSIF bStart THEN                                                    // 出口 2：新批次请求 / New batch requested
        _eState := E_DL_SmxState.eFill;
    END_IF

E_DL_SmxState.eFault:
    ;                                                                     // 故障相：仅段 5 复位沿可迁出 / Only the reset edge leaves this phase

ELSE
    _uFault := 16#0005_03A6;                                             // 故障级：非法相位兜底（归并总码） / Illegal-phase fallback
    _bFault := TRUE;
    bError  := TRUE;
    _eCause := E_DL_SmxCause.ePhaseBad;                                  // 归因：非法相位 / Cause: illegal phase
    _eState := E_DL_SmxState.eFault;

END_CASE

(* —— 段 7：出口单点映射（名实同源；锁存码回放；故障相命令全落） —— *)
IF _bFault THEN
    bInletValveCmd     := FALSE;                                         // 故障相：进料阀关 / Inlet valve closed in fault
    bStirrerFastCmd    := FALSE;                                         // 故障相：高速搅拌停 / High-speed stirrer off in fault
    bVacPumpCmd        := FALSE;                                         // 故障相：真空泵停 / Vacuum pump off in fault
    bDischargeValveCmd := FALSE;                                         // 故障相：出料阀关（安全侧不动料） / Discharge valve closed in fault
    bCycleDone         := FALSE;                                         // 故障相不宣称完成 / No completion claim in fault
ELSE
    bInletValveCmd     := (_eState = E_DL_SmxState.eFill);               // 进料阀仅加料相开 / Inlet open only while filling
    bStirrerFastCmd    := (_eState = E_DL_SmxState.eDisperse);           // 高速搅拌仅分散相开 / Fast stirrer only while dispersing
    bVacPumpCmd        := (_eState = E_DL_SmxState.eDeair);              // 真空泵仅脱泡相开 / Vacuum pump only while de-airing
    bDischargeValveCmd := (_eState = E_DL_SmxState.eDischarge);          // 出料阀仅出料相开 / Discharge valve only while discharging
END_IF
IF _bFault THEN
    nErrId := _uFault;                                                   // 故障锁存码回放 / Replay latched fault code
ELSE
    nErrId := _uInfo;                                                    // 信息码 / Info code
END_IF
bError := _bFault;                                                       // 故障标志与锁存同源（名实双出口，R191） / Flag from latch
eState := _eState;                                                       // 状态出口 / State outlet
eCause := _eCause;                                                       // 成因出口 / Cause outlet

END_FUNCTION_BLOCK
